(* PLC project g_tof_hold, Anonymous Benchmark Suite 1.0 *)
(* stored: creationDateTime 2026-08-26T00:00:00 *)

PROGRAM g_tof_hold
  VAR_INPUT
    Pir : BOOL;
    Button : BOOL;
  END_VAR
  VAR_OUTPUT
    Light : BOOL;
  END_VAR
  VAR
    TOF0 : TOF;
  END_VAR

(* LD diagram, written out as Structured Text *)
TOF0(IN := Pir, PT := T#50ms);
Light := TOF0.Q OR Button;
END_PROGRAM

CONFIGURATION Config0
  RESOURCE Res0 ON PLC
    TASK tcyclic(INTERVAL := T#10ms, PRIORITY := 0);
    PROGRAM inst0 WITH tcyclic : g_tof_hold;
  END_RESOURCE
END_CONFIGURATION
